FUNCTION_BLOCK F (* Negative C1: a second waiting state, but START is only ever left once *)
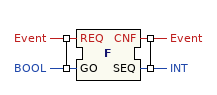
  EVENT_INPUT
    REQ WITH GO;
  END_EVENT
  EVENT_OUTPUT
    CNF WITH SEQ;
  END_EVENT
  VAR_INPUT
    GO : BOOL;
  END_VAR
  VAR_OUTPUT
    SEQ : INT;
  END_VAR
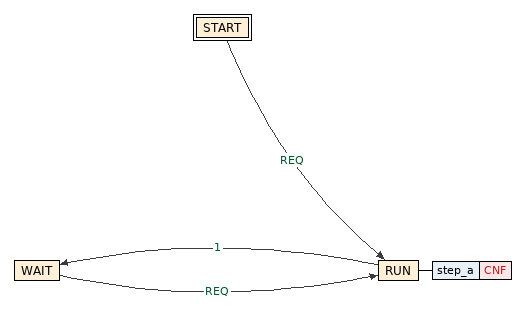
  EC_STATES
    START;
    RUN : step_a -> CNF;
    WAIT;
  END_STATES
  EC_TRANSITIONS
    START TO RUN := REQ;
    RUN TO WAIT := 1;
    WAIT TO RUN := REQ;
  END_TRANSITIONS
  ALGORITHM step_a IN ST:
SEQ := 0;
IF GO THEN
  SEQ := 1;
END_IF;
  END_ALGORITHM
END_FUNCTION_BLOCK
